// TIA Portal V21 export
// export: Created 2000-01-01T00:00:00.0000000Z, ExportSetting None
TYPE "UDT_HMI_MotorRevCtrl"
   STRUCT
      bManualMode { ExternalWritable := 'False'} : Bool;   // HMI手自动切换（TRUE手动）
      bManualFwdCmd { ExternalWritable := 'False'} : Bool;   // HMI手动正转点动/启动
      bManualRevCmd { ExternalWritable := 'False'} : Bool;   // HMI手动反转点动/启动
      bManualStopCmd { ExternalWritable := 'False'} : Bool;   // HMI手动停止
      bResetCmd { ExternalWritable := 'False'} : Bool;   // HMI故障复位命令
      tFeedbackTimeout { ExternalWritable := 'False'} : Time;   // 接触器吸合反馈超时时间（默认 T#2s）
      tReverseDeadband { ExternalWritable := 'False'} : Time;   // 正反转切换停机死区时间（默认 T#1s）
      bRunningFwd { ExternalWritable := 'False'} : Bool;   // 状态反馈：正在正转
      bRunningRev { ExternalWritable := 'False'} : Bool;   // 状态反馈：正在反转
      bFault { ExternalWritable := 'False'} : Bool;   // 状态反馈：综合故障
      wStatus { ExternalWritable := 'False'} : Word;   // 状态码：16#0000正常, 16#8401热过载, 16#8402接触器反馈超时, 16#8403急停激活
   END_STRUCT;
END_TYPE
